(* CODESYS project stringtools.library
   Company: KOSTAL GmbH & Co.KG
   DefaultNamespace: KOSTAL.AF2024.Core.StringTools
   Version: 1.0.0.0
   Placeholder: KOSTAL.AF2024.Core.StringTools
   Author: Frank Dümpelmann
   Description: WSTRING Tools
   Title: KOSTAL.AF2024.Core.StringTools

Project tree, tasks and I/O mapping:
  libraries: KOSTAL.AF2024.Core.ListOf, 1.0.0.0 (KOSTAL GmbH & Co.KG); KOSTAL.AF2024.Core.Settings, 1.0.0.0 (KOSTAL GmbH & Co.KG); KOSTAL.AF2024.Core.System, 1.0.0.0 (KOSTAL GmbH & Co.KG); Tc2_Standard, 3.3.3.0 (Beckhoff Automation GmbH); Tc2_Utilities, 3.4.8.0 (Beckhoff Automation GmbH)
  Enum/
    data type E_ALIGNMENT
  Project Information/
    function F_GetCompany [ST]
    function F_GetTitle [ST]
    function F_GetVersion [ST]
  UTF8/
    CONCAT_UTF8/
      function block FB_Concat_UTF8 [ST]: _clear, addContent, Clear, getResult, FB_exit, FB_init
    Split_UTF8/
      function block FB_Split_UTF8 [ST]: _clear, _execute, Clear, Delimiter, Results, Split, Split_Delimiter, FB_exit, FB_init
      interface I_Split_UTF8: Delimiter, Results
      interface I_Split_UTF8_Owner: Clear, Delimiter, Split, Split_Delimiter
    function F_FLOAT_TO_STRING_UTF8 [ST]
    function F_FormatMask_UTF8 [ST]
    function F_FormatNoMask_UTF8 [ST]
    function F_LREAL_TO_STRING_UTF8 [ST]
    function F_REAL_TO_STRING_UTF8 [ST]
    function F_Replace_UTF8 [ST]
    function F_ToLCase_UTF8 [ST]
    function F_ToUCase_UTF8 [ST]
    function block FB_UrlEscape_UTF8 [ST]: Escape
  Version/
    global variables Global_Version
  WSTRING/
    CONCAT/
      function block FB_Concat [ST]: _clear, addContent, Clear, getResult, FB_exit, FB_init
    SPLIT/
      function block FB_Split [ST]: _clear, _execute, Clear, Delimiter, Results, Split, Split_Delimiter, FB_exit, FB_init
      interface I_Split: Delimiter, Results
      interface I_Split_Owner: Clear, Delimiter, Split, Split_Delimiter
    function F_Replace [ST]
  global variables GVL_CONSTANT
*)

// Enum/E_ALIGNMENT
TYPE E_ALIGNMENT :
	(
		LEFT 	:= 0,
		RIGHT	:= 1,
		CENTER	:= 2
	);
END_TYPE

// Version/Global_Version
{attribute 'TcGenerated'}
{attribute 'no-analysis'}
{attribute 'linkalways'}
// This function has been automatically generated from the project information.
VAR_GLOBAL CONSTANT
	{attribute 'const_non_replaced'}
	stLibVersion_KOSTAL_AF2024_Core_StringTools : ST_LibVersion := (iMajor := 1, iMinor := 0, iBuild := 0, iRevision := 0, nFlags := 0, sVersion := '1.0.0.0');
END_VAR

// GVL_CONSTANT
{attribute 'qualified_only'}
VAR_GLOBAL CONSTANT
	
	OVERFLOW_UTF8	: KOSTAL_AF2024_Core_Settings.T_MaxString_UTF8:= 'OVERFLOW';

	OVERFLOW			: KOSTAL_AF2024_Core_Settings.T_MaxString:= "OVERFLOW";
	
END_VAR

// Project Information/F_GetCompany
// This function has been automatically generated from the project information.
{attribute 'signature_flag' := '1073741824'}
{attribute 'TcGenerated'}
{attribute 'no-analysis'}
FUNCTION F_GetCompany : WSTRING
VAR_INPUT
	
END_VAR

F_GetCompany := "KOSTAL GmbH & Co.KG";

END_FUNCTION

// Project Information/F_GetTitle
// This function has been automatically generated from the project information.
{attribute 'signature_flag' := '1073741824'}
{attribute 'TcGenerated'}
{attribute 'no-analysis'}
FUNCTION F_GetTitle : WSTRING
VAR_INPUT
	
END_VAR

F_GetTitle := "KOSTAL.AF2024.Core.StringTools";

END_FUNCTION

// Project Information/F_GetVersion
// This function has been automatically generated from the project information.
{attribute 'signature_flag' := '1073741824'}
{attribute 'TcGenerated'}
{attribute 'no-analysis'}
FUNCTION F_GetVersion : ST_LibVersion
VAR_INPUT
	
END_VAR

F_GetVersion.iMajor := 1;
F_GetVersion.iMinor := 0;
F_GetVersion.iBuild := 0;
F_GetVersion.iRevision := 0;
F_GetVersion.sVersion := '1.0.0.0';
F_GetVersion.nFlags := 0;

END_FUNCTION

// UTF8/CONCAT_UTF8/FB_Concat_UTF8
FUNCTION_BLOCK PUBLIC FB_Concat_UTF8
VAR
	_List	: KOSTAL_AF2024_Core_listOf.FB_ListOfString_UTF8;
END_VAR

METHOD PROTECTED _clear
VAR_INPUT
END_VAR

_List.clear();
END_METHOD

METHOD PUBLIC addContent : BOOL
VAR_INPUT
	Text	: KOSTAL_AF2024_Core_Settings.T_MaxString_UTF8;
END_VAR

IF _List.NumberOfLines >= _List.maxLine THEN RETURN;	END_IF

addContent:= _List.addLine(Text);
END_METHOD

METHOD PUBLIC Clear
VAR_INPUT
END_VAR

_List.clear();
END_METHOD

METHOD PUBLIC getResult : KOSTAL_AF2024_Core_Settings.T_MaxString_UTF8
VAR_INPUT
END_VAR

VAR
	_udi: UDINT;
END_VAR

getResult:= '';

FOR _udi:= 1 TO _List.NumberOfLines DO
	getResult:= Tc2_Standard.CONCAT(getResult, _List.line_GET(_udi));
END_FOR
END_METHOD

METHOD FB_exit : BOOL
VAR_INPUT
	bInCopyCode : BOOL; // if TRUE, the exit method is called for exiting an instance that is copied afterwards (online change).
END_VAR

_clear();
END_METHOD

METHOD FB_init : BOOL
VAR_INPUT
	bInitRetains : BOOL; // if TRUE, the retain variables are initialized (warm start / cold start)
	bInCopyCode : BOOL;  // if TRUE, the instance afterwards gets moved into the copy code (online change)
END_VAR

_clear();
END_METHOD

END_FUNCTION_BLOCK

// UTF8/Split_UTF8/FB_Split_UTF8
FUNCTION_BLOCK PUBLIC FB_Split_UTF8 IMPLEMENTS I_Split_UTF8, I_Split_UTF8_Owner

VAR
	_CList			: KOSTAL_AF2024_Core_ListOf.FB_ListOfString_UTF8;	//ComponentList
	_Line				: KOSTAL_AF2024_Core_Settings.T_MaxString_UTF8;	
	_delimiter	: STRING(1):= '\';	//default
END_VAR

METHOD PROTECTED _clear
VAR_INPUT
END_VAR

_CList.clear();
_Line				:= '';	
_delimiter	:= '';
END_METHOD

METHOD PROTECTED _execute : BOOL

VAR
	_pos	: INT;
	_work	: KOSTAL_AF2024_Core_Settings.T_MaxString_UTF8;
	_part	: KOSTAL_AF2024_Core_Settings.T_MaxString_UTF8;
END_VAR
_CList.clear();


IF _Line = '' 			THEN	RETURN;	END_IF
IF _delimiter = ''	THEN	RETURN;	END_IF

_work:= _Line;

REPEAT
	
	_pos:= Tc2_Standard.FIND(_work, _delimiter);

	IF _pos > 0 THEN

		IF _pos > 1 THEN	
			_part:= Tc2_Standard.LEFT(_work, _pos - 1);
			_CList.addLine(_part);	
		END_IF

		_work:= Tc2_Standard.RIGHT(_work, Tc2_Standard.LEN(_work) - _pos);
		
	END_IF

UNTIL	(_pos <= 0) OR _CList.NumberOfLines > 255
END_REPEAT

IF _work <> '' THEN _CList.addLine(_work);	END_IF

_execute:= TRUE;
END_METHOD

METHOD PUBLIC Clear
VAR_INPUT
END_VAR

_clear();
END_METHOD

PROPERTY PUBLIC Delimiter : STRING(1)
GET

Delimiter:= _delimiter;
END_GET
SET

_delimiter:= Delimiter;
END_SET
END_PROPERTY

PROPERTY PUBLIC Results : KOSTAL_AF2024_Core_ListOf.I_ListOfString_UTF8
GET

Results:= _CList;
END_GET
END_PROPERTY

METHOD PUBLIC Split : BOOL
VAR_INPUT
	Line	: KOSTAL_AF2024_Core_Settings.T_MaxString_UTF8;
END_VAR
_Line:= Line;

Split:= _execute();
END_METHOD

METHOD PUBLIC Split_Delimiter : BOOL
VAR_INPUT
	Line			: KOSTAL_AF2024_Core_Settings.T_MaxString_UTF8;
	Delimiter	:	STRING(1);
END_VAR
_Line:= Line;

_delimiter:= Delimiter;

Split_Delimiter:= _execute();
END_METHOD

METHOD FB_exit : BOOL
VAR_INPUT
	bInCopyCode : BOOL; // if TRUE, the exit method is called for exiting an instance that is copied afterwards (online change).
END_VAR

_clear();
END_METHOD

METHOD FB_init : BOOL
VAR_INPUT
	bInitRetains : BOOL; // if TRUE, the retain variables are initialized (warm start / cold start)
	bInCopyCode : BOOL;  // if TRUE, the instance afterwards gets moved into the copy code (online change)
END_VAR

_clear();
END_METHOD

END_FUNCTION_BLOCK

// UTF8/Split_UTF8/I_Split_UTF8
INTERFACE I_Split_UTF8 EXTENDS KOSTAL_AF2024_Core_System.I_Interface

PROPERTY PUBLIC Delimiter : STRING(1)
GET
END_GET
END_PROPERTY

PROPERTY PUBLIC Results : KOSTAL_AF2024_Core_ListOf.I_ListOfString_UTF8
GET
END_GET
END_PROPERTY

END_INTERFACE

// UTF8/Split_UTF8/I_Split_UTF8_Owner
INTERFACE I_Split_UTF8_Owner EXTENDS I_Split_UTF8

METHOD PUBLIC Clear
VAR_INPUT
END_VAR
END_METHOD

PROPERTY PUBLIC Delimiter : STRING(1)
SET
END_SET
END_PROPERTY

METHOD PUBLIC Split : BOOL
VAR_INPUT
	Line	: KOSTAL_AF2024_Core_Settings.T_MaxString_UTF8;
END_VAR
END_METHOD

METHOD PUBLIC Split_Delimiter : BOOL
VAR_INPUT
	Line		: KOSTAL_AF2024_Core_Settings.T_MaxString_UTF8;
	Delimiter	:	STRING(1);
END_VAR
END_METHOD

END_INTERFACE

// UTF8/F_FLOAT_TO_STRING_UTF8
(*
Supported Data Types:
REAL;LREAL
*)

FUNCTION F_FLOAT_TO_STRING_UTF8 : STRING(512)

VAR_INPUT
	IN			: Tc2_Utilities.FLOAT;
	Digits	: INT;	//Number of digits after the decimal point
END_VAR

VAR
	_IN			: LREAL;
END_VAR


_IN:= IN;

IF NOT Tc2_Utilities.LrealIsFinite(_IN) THEN	
	F_FLOAT_TO_STRING_UTF8:= GVL_CONSTANT.OVERFLOW_UTF8;
	RETURN;	
ELSIF Tc2_Utilities.LrealIsNaN(_IN) THEN	
	F_FLOAT_TO_STRING_UTF8:= GVL_CONSTANT.OVERFLOW_UTF8;
	RETURN;	
END_IF

F_FLOAT_TO_STRING_UTF8:= Tc2_Utilities.LREAL_TO_FMTSTR(IN, Digits, FALSE);

END_FUNCTION

// UTF8/F_FormatMask_UTF8
(*

:Author: Frank Dümpelmann <f.duempelmann@kostal.com>, Martin Hundt <m.hundt@kostal.com>
:Date: 2018-10-29

Function
========
| Formats =line= to the length of =mask= with the characters defined in =mask= and given =alignment=
| If =line= is longer than =mask=, the method will return =line= with the original length

Methods and Properties
======================
| line	: STRING(255) - String to format
| mask	: STRING(255) - e.g., '00000' formats line to 5 characters, filling up with the placeholder 0 
| alignment	: E_ALIGNMENT - Alignment of the original string

Usage sample:
=============

.. code:: 

	PROGRAM MAIN
	VAR	
		_Test : STRING(255) := 'test';
	END_VAR
	
	_Test := F_Format(line := _Test, mask:= 'xxxxxxxxxx', alignment:=E_ALIGNMENT.Left);

*)


FUNCTION F_FormatMask_UTF8 : KOSTAL_AF2024_Core_Settings.T_MaxString_UTF8
VAR_INPUT
	line	: KOSTAL_AF2024_Core_Settings.T_MaxString_UTF8;	//
	mask	: KOSTAL_AF2024_Core_Settings.T_MaxString_UTF8;			//f.a. '00000' defines the minimum lenght and placeholder for empty string position 
	alignment	: E_ALIGNMENT;
END_VAR
VAR
END_VAR


IF alignment = E_ALIGNMENT.LEFT THEN

	IF Tc2_Standard.LEN(mask) > Tc2_Standard.LEN(line) THEN
		F_FormatMask_UTF8:= Tc2_Standard.LEFT(Tc2_Standard.CONCAT(line, mask), Tc2_Standard.LEN(mask));		
	ELSE
		F_FormatMask_UTF8:= Tc2_Standard.LEFT(Tc2_Standard.CONCAT(line, mask), Tc2_Standard.LEN(line));		
	END_IF
	
ELSIF alignment = E_ALIGNMENT.RIGHT THEN

	IF Tc2_Standard.LEN(mask) > Tc2_Standard.LEN(line) THEN
		F_FormatMask_UTF8:= Tc2_Standard.RIGHT(Tc2_Standard.CONCAT(mask, line), Tc2_Standard.LEN(mask));		
	ELSE
		F_FormatMask_UTF8:= Tc2_Standard.RIGHT(Tc2_Standard.CONCAT(mask, line), Tc2_Standard.LEN(line));		
	END_IF

ELSE
	F_FormatMask_UTF8:= '';		
END_IF

END_FUNCTION

// UTF8/F_FormatNoMask_UTF8
(*

:Author: Martin Hundt <m.hundt@kostal.com>
:Date: 2021-12-10

Function
========
| Formats =line= to the length of =formatLength= with the characters =char= and given =alignment=
| If =line= is longer than =formatLength=, the method will return =line= with the original length

Methods and Properties
======================
| line			: STRING(255) - String to format
| formatLength	: UINT - length of formatted string 
| char			: STRING(1) - Character to fill the sting. Default: Space 
| alignment		: E_ALIGNMENT - Alignment of the return string

Usage sample:
=============
See best practice
*)


FUNCTION F_FormatNoMask_UTF8 : KOSTAL_AF2024_Core_Settings.T_MaxString_UTF8
VAR_INPUT
	line					: KOSTAL_AF2024_Core_Settings.T_MaxString_UTF8;	//
	formatLength	: UINT;
	char					: STRING(1); 
	alignment			: E_ALIGNMENT;
END_VAR
VAR
	_stringLength	: UINT;
	_fillLength		: UINT;
	_out					: KOSTAL_AF2024_Core_Settings.T_MaxString_UTF8;
	_i						: UINT;
END_VAR

IF char = '' THEN 
	char := ' '; 
END_IF
_stringLength := INT_TO_UINT(Tc2_Standard.LEN(line));

IF _stringLength >= formatLength THEN
	_out := line;
ELSIF alignment = E_ALIGNMENT.LEFT THEN
	_out := line;
	FOR _i:= _stringLength TO formatLength DO
		_out := Tc2_Standard.CONCAT(_out, char);
	END_FOR

	
ELSIF alignment = E_ALIGNMENT.RIGHT THEN
	
	FOR _i:= 1 TO (formatLength - _stringLength) DO
		_out := Tc2_Standard.CONCAT(_out, char);
	END_FOR
	_out := Tc2_Standard.CONCAT(_out, line);
	
ELSIF alignment = E_ALIGNMENT.CENTER THEN	
	
	_fillLength := (formatLength-_stringLength)/2;
	
	FOR _i:=0 TO formatLength DO	//Fill with spaces
		_out := CONCAT(_out, char);
	END_FOR
	
	
	_out :=  Tc2_Standard.INSERT(_out, line,_fillLength + 1);
		
END_IF

F_FormatNoMask_UTF8:= _out;

END_FUNCTION

// UTF8/F_LREAL_TO_STRING_UTF8
(*
Supported Data Types:
REAL;LREAL
*)

FUNCTION F_LREAL_TO_STRING_UTF8 : STRING(512)

VAR_INPUT
	IN			: LREAL;
	Digits	: INT;	//Number of digits after the decimal point
END_VAR

VAR
	_IN			: LREAL;
END_VAR

_IN:= IN;

IF NOT Tc2_Utilities.LrealIsFinite(_IN) THEN	
	F_LREAL_TO_STRING_UTF8:= GVL_CONSTANT.OVERFLOW_UTF8;
	RETURN;	
ELSIF Tc2_Utilities.LrealIsNaN(_IN) THEN	
	F_LREAL_TO_STRING_UTF8:= GVL_CONSTANT.OVERFLOW_UTF8;
	RETURN;	
END_IF

F_LREAL_TO_STRING_UTF8:= Tc2_Utilities.LREAL_TO_FMTSTR(IN, Digits, FALSE);

END_FUNCTION

// UTF8/F_REAL_TO_STRING_UTF8
(*
Supported Data Types:
REAL;LREAL
*)
FUNCTION F_REAL_TO_STRING_UTF8 : STRING(512)

VAR_INPUT
	IN			: REAL;
	Digits	: INT;	//Number of digits after the decimal point
END_VAR

VAR
	_T_Arg: Tc2_Utilities.T_Arg;
END_VAR


_T_Arg:= Tc2_Utilities.F_REAL(IN);

IF NOT Tc2_Utilities.IsFinite(_T_Arg) THEN	
	F_REAL_TO_STRING_UTF8:= GVL_CONSTANT.OVERFLOW_UTF8;
	RETURN;	
END_IF

F_REAL_TO_STRING_UTF8:= Tc2_Utilities.LREAL_TO_FMTSTR(IN, Digits, FALSE);

END_FUNCTION

// UTF8/F_Replace_UTF8
(*

:Author: Frank Dümpelmann <f.duempelmann@kostal.com>, Martin Hundt <m.hundt@kostal.com>
:Date: 2018-10-30

Function
========
Replace all occurencies of a given string with another string

Methods and Properties
======================
| source 						: KOSTAL_TC3_Core_Settings.T_MaxString - string to replace in
| toReplace					: KOSTAL_TC3_Core_Settings.T_MaxString - string to replace
| replaceWith 			: KOSTAL_TC3_Core_Settings.T_MaxString - string to replace with
| numberOfReplaces	: Replace only the first X occurencies from left (default: -1, replace all occurrencies)

*) 

FUNCTION F_Replace_UTF8 : KOSTAL_AF2024_Core_Settings.T_MaxString_UTF8

VAR_INPUT
	source						: KOSTAL_AF2024_Core_Settings.T_MaxString_UTF8;
	toReplace					: KOSTAL_AF2024_Core_Settings.T_MaxString_UTF8;
	replaceWith				: KOSTAL_AF2024_Core_Settings.T_MaxString_UTF8;
	numberOfReplaces	: INT:= -1;	(*INT:= -1 defines to replace all occurrences *)
END_VAR

VAR
	_index				: INT;
	_pos					: INT;
	_replaced			: KOSTAL_AF2024_Core_Settings.T_MaxString_UTF8;
	_toReplaceLen	: INT;
	_searchPos		: INT;
	_searchString	: KOSTAL_AF2024_Core_Settings.T_MaxString_UTF8;
	_i: INT;
END_VAR

IF 		numberOfReplaces  =  0  									THEN	F_Replace_UTF8:= source;	RETURN;	//no replacement required
ELSIF Tc2_Standard.FIND(source, toReplace) = 0	THEN 	F_Replace_UTF8:= source;	RETURN;	//no replacement required
ELSIF numberOfReplaces  <  0  									THEN	_index:= LEN(source);				//full replacement required
ELSE																									_index:= numberOfReplaces;	//replacement limmitted by numberOfReplaces
END_IF

//prepare
_replaced			:= '';
_toReplaceLen	:= Tc2_Standard.LEN(toReplace);
_searchString	:= source;
_searchPos		:= 1;


FOR _i:= 1 TO _index DO
	
	//find next to replace content
	_pos:= Tc2_Standard.FIND(_searchString, toReplace);

	//no further to replace found
	IF _pos = 0 THEN	EXIT;	END_IF
		
	//get left n characters until _pos
	IF _pos > 1 THEN	_replaced:= Tc2_Standard.CONCAT(_replaced, Tc2_Standard.LEFT(_searchString, _pos - 1));	END_IF

	//add replaced content
	_replaced:= Tc2_Standard.CONCAT(_replaced, replaceWith);
	
	//Capture the remaining characters to be checked   
	_searchString:= Tc2_Standard.RIGHT(_searchString, Tc2_Standard.LEN(_searchString) - (_pos - 1) - _toReplaceLen);
	
END_FOR

_replaced:= Tc2_Standard.CONCAT(_replaced, _searchString);
 	
F_Replace_UTF8:= _replaced;

END_FUNCTION

// UTF8/F_ToLCase_UTF8
(*

:Author: Frank Dümpelmann <f.duempelmann@kostal.com>, Martin Hundt <m.hundt@kostal.com>
:Date: 2018-10-30

Function
========
Set all characters in the string to upper case

Usage notes
===============
| Only ASCII charset is supported

*) 

FUNCTION F_ToLCase_UTF8 : KOSTAL_AF2024_Core_Settings.T_MaxString_UTF8

VAR_INPUT
	IN		: KOSTAL_AF2024_Core_Settings.T_MaxString_UTF8;
END_VAR

VAR
	_pos		: INT;
	_sign	: STRING(1);
END_VAR


F_ToLCase_UTF8:= Tc2_Utilities.F_ToLCase(IN);

END_FUNCTION

// UTF8/F_ToUCase_UTF8
(*

:Author: Frank Dümpelmann <f.duempelmann@kostal.com>, Martin Hundt <m.hundt@kostal.com>
:Date: 2018-10-30

Function
========
Set all characters in the string to upper case

Usage notes
===============
| Only ASCII charset is supported

*) 

FUNCTION F_ToUCase_UTF8 : KOSTAL_AF2024_Core_Settings.T_MaxString_UTF8

VAR_INPUT
	IN		: KOSTAL_AF2024_Core_Settings.T_MaxString_UTF8;
END_VAR

VAR
	_pos		: INT;
	_sign	: STRING(1);
END_VAR


F_ToUCase_UTF8:= Tc2_Utilities.F_ToUCase(IN);

END_FUNCTION

// UTF8/FB_UrlEscape_UTF8
(*

:Author: Frank Dümpelmann <f.duempelmann@kostal.com>
:Date: 2018-10-30

Function
========
Class for replacing invalid characters in a URL with escape sequences. 
*)

FUNCTION_BLOCK PUBLIC FB_UrlEscape_UTF8

VAR
	_s	: KOSTAL_AF2024_Core_Settings.T_MaxString_UTF8;
END_VAR

(*
Return TRUE 	: At least one character was escaped.
Return FALSE	: No character was escaped.
*)
METHOD PUBLIC Escape : BOOL

VAR_INPUT
	URL					: KOSTAL_AF2024_Core_Settings.T_MaxString_UTF8;
	URL_Escaped	: REFERENCE TO KOSTAL_AF2024_Core_Settings.T_MaxString_UTF8;	//Reference to a resultstring
END_VAR
//$24 (Hex) is ASCII Code for %

_s:= URL;

IF _s <> '' THEN

	_s:= F_Replace_UTF8(_s,'%', '%25', -1);	
	
	_s:= F_Replace_UTF8(_s,' ', '%20', -1);
	_s:= F_Replace_UTF8(_s,'<', '%3C', -1);
	_s:= F_Replace_UTF8(_s,'>', '%3E', -1);
	_s:= F_Replace_UTF8(_s,'#', '%23', -1);
	_s:= F_Replace_UTF8(_s,'+', '%2B', -1);
	_s:= F_Replace_UTF8(_s,'{', '%7B', -1);
	_s:= F_Replace_UTF8(_s,'}', '%7D', -1);
	_s:= F_Replace_UTF8(_s,'|', '%7C', -1);
	_s:= F_Replace_UTF8(_s,'\', '%5C', -1);
	_s:= F_Replace_UTF8(_s,'^', '%5E', -1);
	_s:= F_Replace_UTF8(_s,'~', '%7E', -1);
	_s:= F_Replace_UTF8(_s,'[', '%5B', -1);
	_s:= F_Replace_UTF8(_s,']', '%5D', -1);
	_s:= F_Replace_UTF8(_s,'$'', '%60', -1);
	_s:= F_Replace_UTF8(_s,';', '%3B', -1);
	_s:= F_Replace_UTF8(_s,'/', '%2F', -1);
	_s:= F_Replace_UTF8(_s,'?', '%3F', -1);
	_s:= F_Replace_UTF8(_s,':', '%3A', -1);
	_s:= F_Replace_UTF8(_s,'@', '%40', -1);
	_s:= F_Replace_UTF8(_s,'=', '%3D', -1);
	_s:= F_Replace_UTF8(_s,'&', '%26', -1);
	_s:= F_Replace_UTF8(_s,'$$', '%24', -1);

END_IF

Escape:= _s <> URL;

IF __ISVALIDREF(URL_Escaped) THEN	URL_Escaped:= _s;	END_IF
END_METHOD

END_FUNCTION_BLOCK

// WSTRING/CONCAT/FB_Concat
FUNCTION_BLOCK PUBLIC FB_Concat
VAR
	_List	: FB_ListOfString;
END_VAR

METHOD PROTECTED _clear
VAR_INPUT
END_VAR

_List.clear();
END_METHOD

METHOD PUBLIC addContent : BOOL
VAR_INPUT
	Text	: KOSTAL_AF2024_Core_Settings.T_MaxString;
END_VAR

IF _List.NumberOfLines >= _List.maxLine THEN RETURN;	END_IF

addContent:= _List.addLine(Text);
END_METHOD

METHOD PUBLIC Clear
VAR_INPUT
END_VAR

_List.clear();
END_METHOD

METHOD PUBLIC getResult : KOSTAL_AF2024_Core_Settings.T_MaxString
VAR_INPUT
END_VAR

VAR
	_udi: UDINT;
END_VAR

getResult:= "";

FOR _udi:= 1 TO _List.NumberOfLines DO
	getResult:= Tc2_Standard.WCONCAT(getResult, _List.line_GET(_udi));
END_FOR
END_METHOD

METHOD FB_exit : BOOL
VAR_INPUT
	bInCopyCode : BOOL; // if TRUE, the exit method is called for exiting an instance that is copied afterwards (online change).
END_VAR

_clear();
END_METHOD

METHOD FB_init : BOOL
VAR_INPUT
	bInitRetains : BOOL; // if TRUE, the retain variables are initialized (warm start / cold start)
	bInCopyCode : BOOL;  // if TRUE, the instance afterwards gets moved into the copy code (online change)
END_VAR

_clear();
END_METHOD

END_FUNCTION_BLOCK

// WSTRING/SPLIT/FB_Split
FUNCTION_BLOCK PUBLIC FB_Split IMPLEMENTS I_Split, I_Split_Owner

VAR
	_CList			: KOSTAL_AF2024_Core_ListOf.FB_ListOfString;	//ComponentList
	_Line				: KOSTAL_AF2024_Core_Settings.T_MaxString;	
	_delimiter	: WSTRING(1):= "\";	//default
END_VAR

METHOD PROTECTED _clear
VAR_INPUT
END_VAR

_CList.clear();
_Line				:= "";	
_delimiter	:= "";
END_METHOD

METHOD PROTECTED _execute : BOOL

VAR
	_pos	: INT;
	_work	: KOSTAL_AF2024_Core_Settings.T_MaxString;
	_part	: KOSTAL_AF2024_Core_Settings.T_MaxString;
END_VAR
_CList.clear();


IF _Line = "" 			THEN	RETURN;	END_IF
IF _delimiter = ""	THEN	RETURN;	END_IF

_work:= _Line;

REPEAT
	
	_pos:= Tc2_Standard.WFIND(_work, _delimiter);

	IF _pos > 0 THEN

		IF _pos > 1 THEN	
			_part:= Tc2_Standard.WLEFT(_work, _pos - 1);
			_CList.addLine(_part);	
		END_IF

		_work:= Tc2_Standard.WRIGHT(_work, Tc2_Standard.WLEN(_work) - _pos);
		
	END_IF

UNTIL	(_pos <= 0) OR _CList.NumberOfLines > 255
END_REPEAT

IF _work <> "" THEN _CList.addLine(_work);	END_IF

_execute:= TRUE;
END_METHOD

METHOD PUBLIC Clear
VAR_INPUT
END_VAR

_clear();
END_METHOD

PROPERTY PUBLIC Delimiter : WSTRING(1)
GET

Delimiter:= _delimiter;
END_GET
SET

_delimiter:= Delimiter;
END_SET
END_PROPERTY

PROPERTY PUBLIC Results : KOSTAL_AF2024_Core_ListOf.I_ListOfString
GET

Results:= _CList;
END_GET
END_PROPERTY

METHOD PUBLIC Split : BOOL
VAR_INPUT
	Line	: KOSTAL_AF2024_Core_Settings.T_MaxString;
END_VAR
_Line:= Line;

Split:= _execute();
END_METHOD

METHOD PUBLIC Split_Delimiter : BOOL
VAR_INPUT
	Line			: KOSTAL_AF2024_Core_Settings.T_MaxString;
	Delimiter	:	WSTRING(1);
END_VAR
_Line:= Line;

_delimiter:= Delimiter;

Split_Delimiter:= _execute();
END_METHOD

METHOD FB_exit : BOOL
VAR_INPUT
	bInCopyCode : BOOL; // if TRUE, the exit method is called for exiting an instance that is copied afterwards (online change).
END_VAR

_clear();
END_METHOD

METHOD FB_init : BOOL
VAR_INPUT
	bInitRetains : BOOL; // if TRUE, the retain variables are initialized (warm start / cold start)
	bInCopyCode : BOOL;  // if TRUE, the instance afterwards gets moved into the copy code (online change)
END_VAR

_clear();
END_METHOD

END_FUNCTION_BLOCK

// WSTRING/SPLIT/I_Split
INTERFACE I_Split EXTENDS KOSTAL_AF2024_Core_System.I_Interface

PROPERTY PUBLIC Delimiter : WSTRING(1)
GET
END_GET
END_PROPERTY

PROPERTY PUBLIC Results : I_ListOfString
GET
END_GET
END_PROPERTY

END_INTERFACE

// WSTRING/SPLIT/I_Split_Owner
INTERFACE I_Split_Owner EXTENDS I_Split

METHOD PUBLIC Clear
VAR_INPUT
END_VAR
END_METHOD

PROPERTY PUBLIC Delimiter : WSTRING(1)
SET
END_SET
END_PROPERTY

METHOD PUBLIC Split : BOOL
VAR_INPUT
	Line	: KOSTAL_AF2024_Core_Settings.T_MaxString;
END_VAR
END_METHOD

METHOD PUBLIC Split_Delimiter : BOOL
VAR_INPUT
	Line			: KOSTAL_AF2024_Core_Settings.T_MaxString;
	Delimiter	:	WSTRING(1);
END_VAR
END_METHOD

END_INTERFACE

// WSTRING/F_Replace
(*

:Author: Frank Dümpelmann <f.duempelmann@kostal.com>, Martin Hundt <m.hundt@kostal.com>
:Date: 2018-10-30

Function
========
Replace all occurencies of a given string with another string

Methods and Properties
======================
| source 						: KOSTAL_TC3_Core_Settings.T_MaxString - string to replace in
| toReplace					: KOSTAL_TC3_Core_Settings.T_MaxString - string to replace
| replaceWith 			: KOSTAL_TC3_Core_Settings.T_MaxString - string to replace with
| numberOfReplaces	: Replace only the first X occurencies from left (default: -1, replace all occurrencies)

*) 

FUNCTION F_Replace : KOSTAL_AF2024_Core_Settings.T_MaxString

VAR_INPUT
	source						: KOSTAL_AF2024_Core_Settings.T_MaxString;
	toReplace					: KOSTAL_AF2024_Core_Settings.T_MaxString;
	replaceWith				: KOSTAL_AF2024_Core_Settings.T_MaxString;
	numberOfReplaces	: INT:= -1;	(*INT:= -1 defines to replace all occurrences *)
END_VAR

VAR
	_index				: INT;
	_pos					: INT;
	_replaced			: KOSTAL_AF2024_Core_Settings.T_MaxString;
	_toReplaceLen	: INT;
	_searchPos		: INT;
	_searchString	: KOSTAL_AF2024_Core_Settings.T_MaxString;
	_i: INT;
END_VAR



IF 		numberOfReplaces  =  0  									THEN	F_Replace:= source;	RETURN;	//no replacement required
ELSIF Tc2_Standard.WFIND(source, toReplace) = 0	THEN 	F_Replace:= source;	RETURN;	//no replacement required
ELSIF numberOfReplaces  <  0  									THEN	_index:= WLEN(source);				//full replacement required
ELSE																									_index:= numberOfReplaces;	//replacement limmitted by numberOfReplaces
END_IF

//prepare
_replaced			:= "";
_toReplaceLen	:= Tc2_Standard.WLEN(toReplace);
_searchString	:= source;
_searchPos		:= 1;


FOR _i:= 1 TO _index DO
	
	//find next to replace content
	_pos:= Tc2_Standard.WFIND(_searchString, toReplace);

	//no further to replace found
	IF _pos = 0 THEN	EXIT;	END_IF
		
	//get left n characters until _pos
	IF _pos > 1 THEN	_replaced:= Tc2_Standard.WCONCAT(_replaced, Tc2_Standard.WLEFT(_searchString, _pos - 1));	END_IF

	//add replaced content
	_replaced:= Tc2_Standard.WCONCAT(_replaced, replaceWith);
	
	//Capture the remaining characters to be checked   
	_searchString:= Tc2_Standard.WRIGHT(_searchString, Tc2_Standard.WLEN(_searchString) - (_pos - 1) - _toReplaceLen);
	
END_FOR

_replaced:= Tc2_Standard.WCONCAT(_replaced, _searchString);
 	
F_Replace:= _replaced;

END_FUNCTION
